(* Logix 5000 project; controller R400_500_XLS vendor 1 type 14 code 216 rev 31.11; software revision 31.01; part 7 of 32 *)
(* tags used below, declared in another part *)
   Abort1 : DINT;   // Not Used
   Abort2 : SINT;
   CURRENT_CYCLE : DINT;
   CycExcBuffer : UDT_CYCLE;
   CycleSequence : UDT_CYCLE_SEQUENCE;
   Drain_RcvryTnk_with_Sump : DINT;   // 0 = Close Recovery Tank Drain Valve 1 = Open Recovery Tank Drain Valve
   DrnSmp : DINT;
   DRYING : DINT;   // Drying id number
   F1rinse : DINT;   // Not Used
   F2rinse : DINT;   // Not Used
   F3rinse : DINT;   // Not Used
   FC65_Enabled_signal : BOOL;   // Enables the treatment evaluation
   FC65_Treatment_counter : DINT;   // Treatment counter
   Fill_Sump : DINT;
   FINALRINSE_1 : DINT;   // Final rinse 1 id number
   FINALRINSE_9 : DINT;   // Final rinse 9 id number
   HeatSmp : DINT;
   Inj_Time : SINT;   // Time based chemical injection steps
   M : DINT[5];   // Memory Bits
   ONS_FC13 : DINT;
   ONS_FC65 : DINT;
   OPR_16_TreatPrint_Ptr : DINT;
   PREWASH_1 : DINT;   // Pre-wash 1 id number
   PREWASH_2 : DINT;   // Pre-wash 2 id number
   PREWASH_3 : DINT;   // Pre-wash 3 id number
   PREWASH_4 : DINT;   // Pre-wash 4 id number
   printCycleParameters : STRING[2];
   PWHeat : SINT;
   Rcvry_Tnk_Tmp : REAL;   // Water Temperature of the Heat Recovery Tank
   RINSE_1 : DINT;   // Rinse 1 id number
   RINSE_2 : DINT;   // Rinse 2 id number
   RINSE_3 : DINT;   // Rinse 3 id number
   RINSE_4 : DINT;   // Rinse 4 id number
   Run : DINT;
   sCRLF : STRING;
   sPrntArray : STRING[300];   // Printer String Array
   SumpWaterVolume : DINT;   // Sump Water Volume 0 =Low 1= High
   Tmr : TIMER[107];
   Trt_Drying : SINT;
   Trt_PrWsh : DINT;
   Trt_Rinse : DINT;   // Rinse steps
   Trt_Wsh : DINT;
   VENTING : DINT;   // Venting id number
   WASH_1 : DINT;   // Wash 1 id number
   WASH_2 : DINT;   // Wash 2 id number
   WASH_3 : DINT;   // Wash 3 id number
   WASH_4 : DINT;   // Wash 4 id number
   WASH_5 : DINT;   // Wash 5 id number
   CycleName : STRING[12];
   EnaDisPrinter : BOOL;   // Screen 80 Enable/Disable Printer button
   msg : BOOL[512];
   Msg_Abort : SINT;
   PrintIndex : DINT;
   Screen_Ctrl : DINT;   // PLC Screen Request
   sDateTime : STRING;   // String Date Time
   Tpb : DINT[11];
   TreatmentPtr : DINT;
   Unit : Hrdwre;   // Unit Configuration
(* MainProgram, continued *)

ROUTINE OPR_15_WSH_13_ABORT   (* ladder *)
// This module manage the abort sequence.
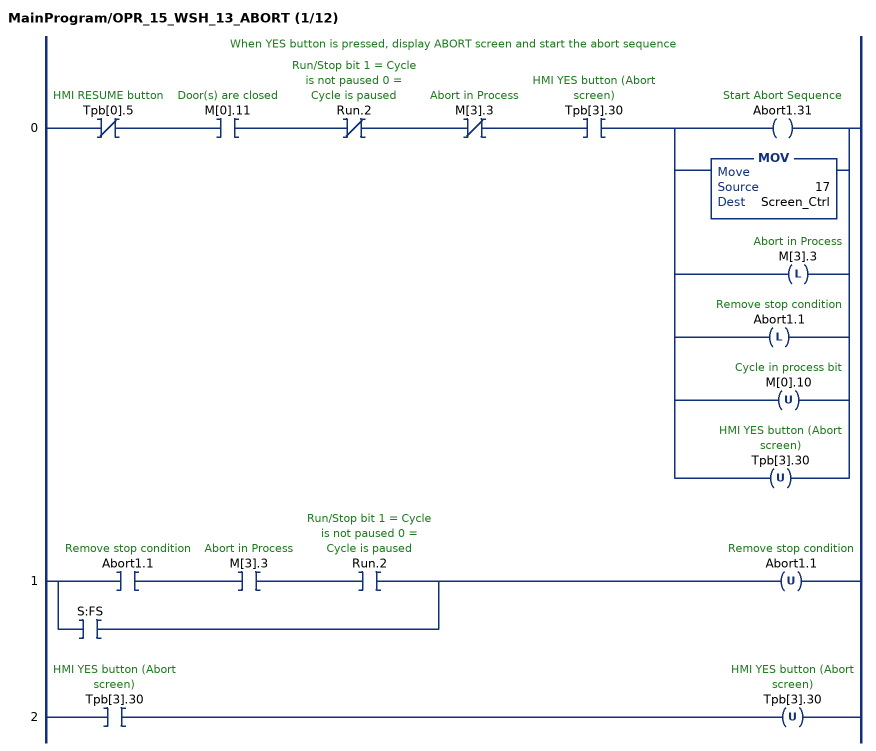
   // When YES button is pressed, display ABORT screen and start the abort sequence
   0: XIO(Tpb[0].5)XIC(M[0].11)XIO(Run.2)XIO(M[3].3)XIC(Tpb[3].30)[OTE(Abort1.31) ,MOV(17,Screen_Ctrl) ,OTL(M[3].3) ,OTL(Abort1.1) ,OTU(M[0].10) ,OTU(Tpb[3].30) ];
   1: [XIC(Abort1.1) XIC(M[3].3) XIC(Run.2) ,XIC(S:FS) ]OTU(Abort1.1);
   2: XIC(Tpb[3].30)OTU(Tpb[3].30);
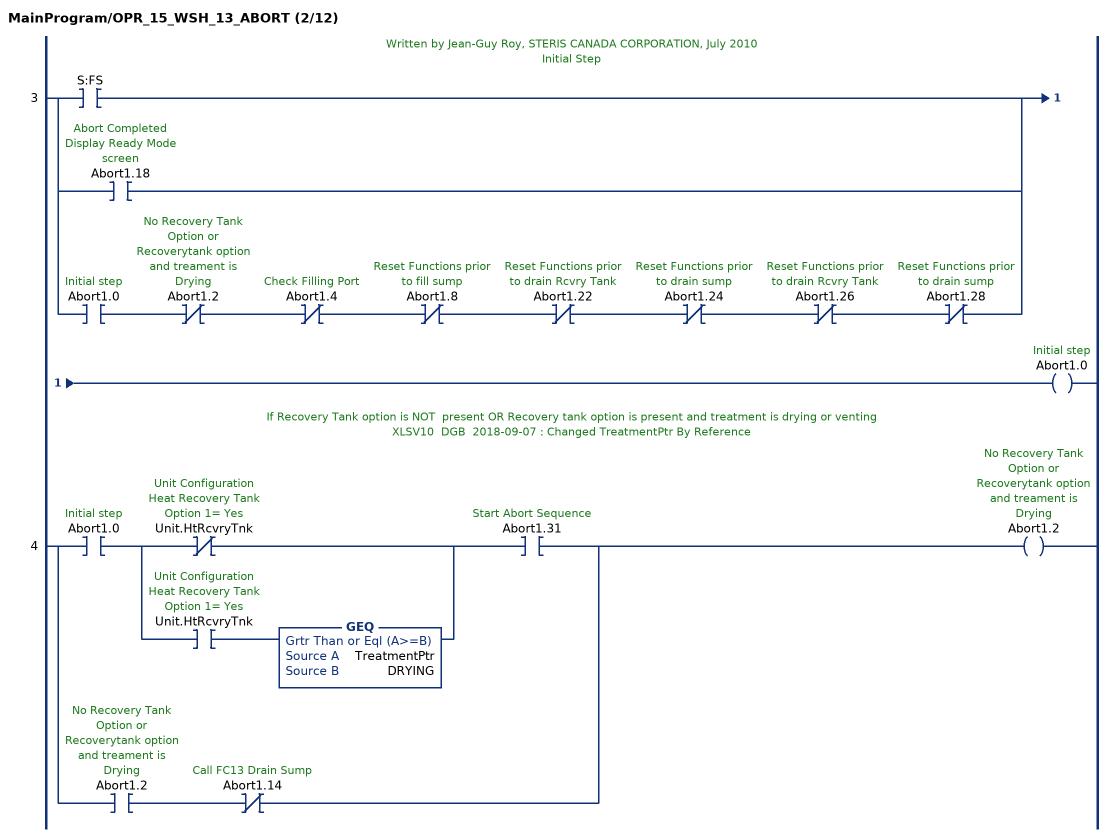
   // Written by Jean-Guy Roy, STERIS CANADA CORPORATION, July 2010
   // Initial Step
   3: [XIC(S:FS) ,XIC(Abort1.18) ,XIC(Abort1.0) XIO(Abort1.2) XIO(Abort1.4) XIO(Abort1.8) XIO(Abort1.22) XIO(Abort1.24) XIO(Abort1.26) XIO(Abort1.28) ]OTE(Abort1.0);
   // If Recovery Tank option is NOT  present OR Recovery tank option is present and treatment is drying or venting
   // XLSV10  DGB  2018-09-07 : Changed TreatmentPtr By Reference
   4: [XIC(Abort1.0) [XIO(Unit.HtRcvryTnk) ,XIC(Unit.HtRcvryTnk) GEQ(TreatmentPtr,DRYING) ] XIC(Abort1.31) ,XIC(Abort1.2) XIO(Abort1.14) ]OTE(Abort1.2);
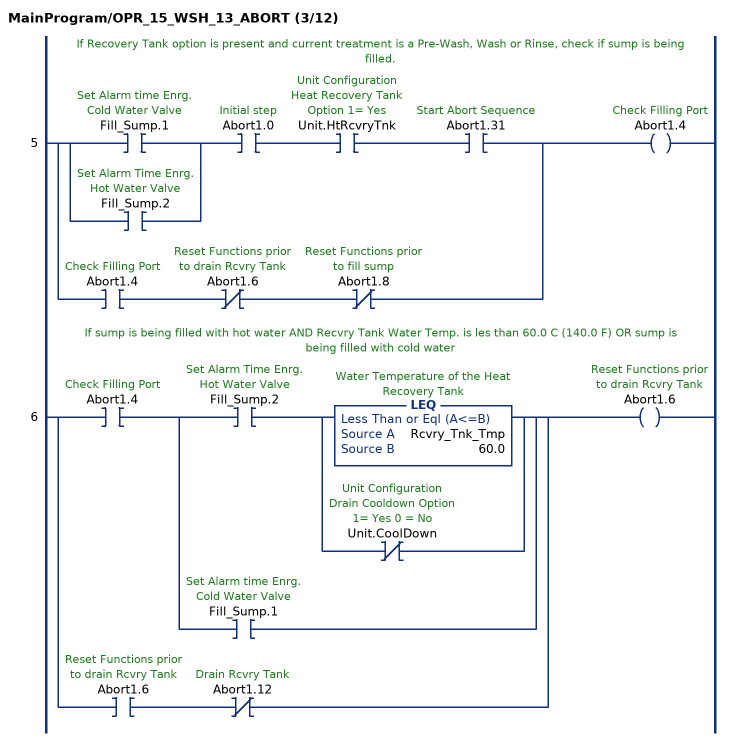
   // If Recovery Tank option is present and current treatment is a Pre-Wash, Wash or Rinse, check if sump is being filled.
   5: [[XIC(Fill_Sump.1) ,XIC(Fill_Sump.2) ] XIC(Abort1.0) XIC(Unit.HtRcvryTnk) XIC(Abort1.31) ,XIC(Abort1.4) XIO(Abort1.6) XIO(Abort1.8) ]OTE(Abort1.4);
   // If sump is being filled with hot water AND Recvry Tank Water Temp. is les than 60.0 C (140.0 F) OR sump is being filled with cold water
   6: [XIC(Abort1.4) [XIC(Fill_Sump.2) [LEQ(Rcvry_Tnk_Tmp,60.0) ,XIO(Unit.CoolDown) ] ,XIC(Fill_Sump.1) ] ,XIC(Abort1.6) XIO(Abort1.12) ]OTE(Abort1.6);
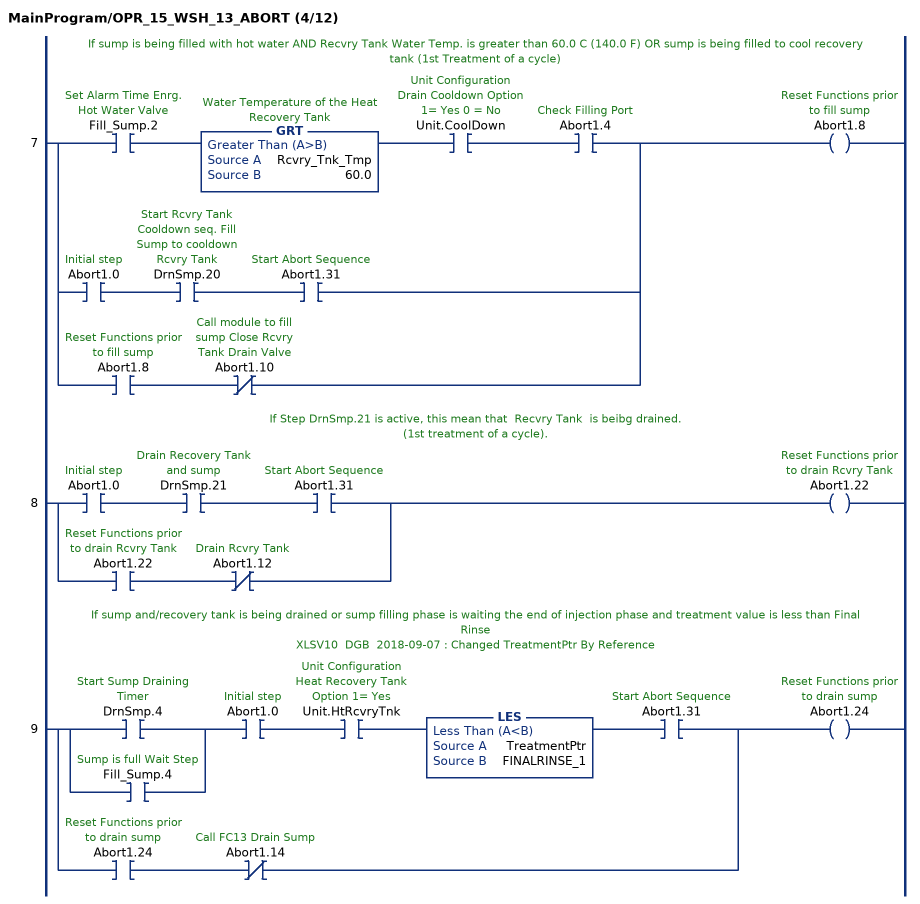
   // If sump is being filled with hot water AND Recvry Tank Water Temp. is greater than 60.0 C (140.0 F) OR sump is being filled to cool recovery tank (1st Treatment of a cycle)
   7: [[XIC(Fill_Sump.2) GRT(Rcvry_Tnk_Tmp,60.0) XIC(Unit.CoolDown) XIC(Abort1.4) ,XIC(Abort1.0) XIC(DrnSmp.20) XIC(Abort1.31) ] ,XIC(Abort1.8) XIO(Abort1.10) ]OTE(Abort1.8);
   // If Step DrnSmp.21 is active, this mean that  Recvry Tank  is beibg drained.
   //  (1st treatment of a cycle).
   8: [XIC(Abort1.0) XIC(DrnSmp.21) XIC(Abort1.31) ,XIC(Abort1.22) XIO(Abort1.12) ]OTE(Abort1.22);
   // If sump and/recovery tank is being drained or sump filling phase is waiting the end of injection phase and treatment value is less than Final Rinse
   // XLSV10  DGB  2018-09-07 : Changed TreatmentPtr By Reference
   9: [[XIC(DrnSmp.4) ,XIC(Fill_Sump.4) ] XIC(Abort1.0) XIC(Unit.HtRcvryTnk) LES(TreatmentPtr,FINALRINSE_1) XIC(Abort1.31) ,XIC(Abort1.24) XIO(Abort1.14) ]OTE(Abort1.24);
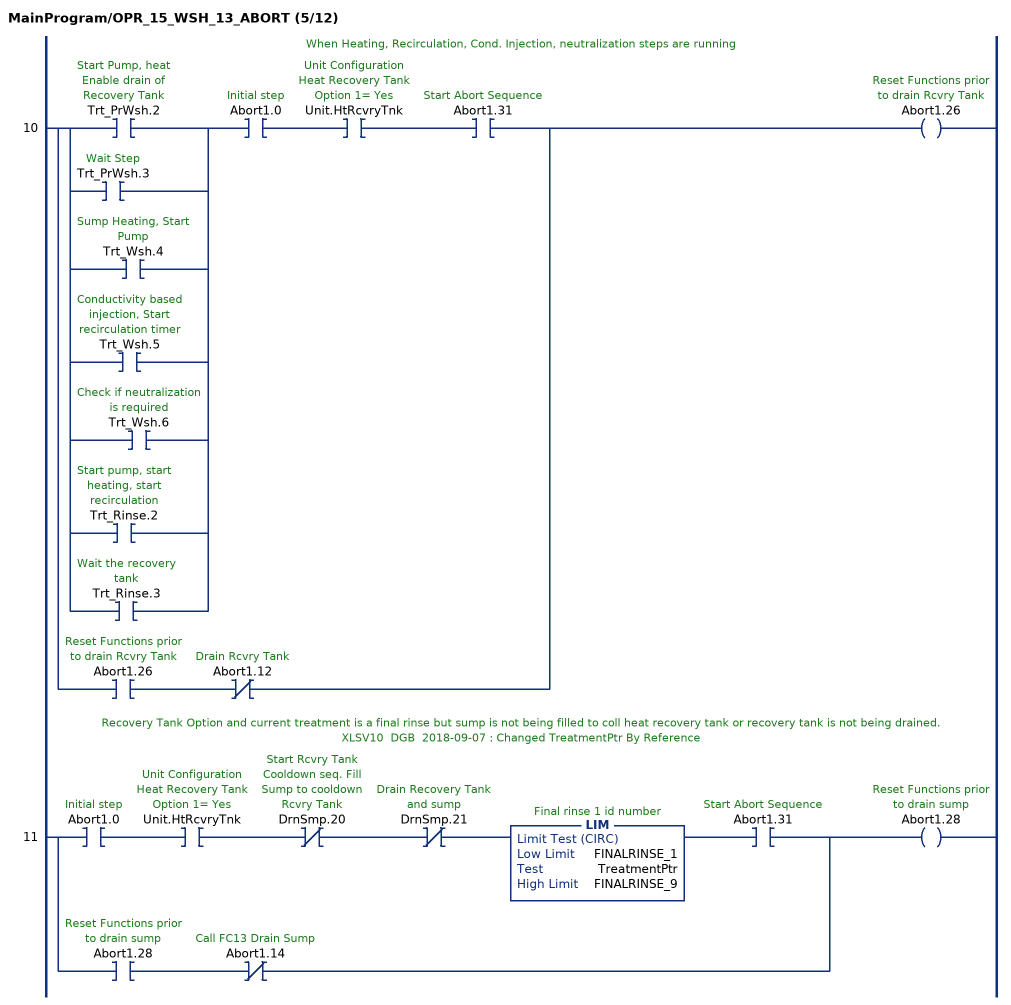
   // When Heating, Recirculation, Cond. Injection, neutralization steps are running
   10: [[XIC(Trt_PrWsh.2) ,XIC(Trt_PrWsh.3) ,XIC(Trt_Wsh.4) ,XIC(Trt_Wsh.5) ,XIC(Trt_Wsh.6) ,XIC(Trt_Rinse.2) ,XIC(Trt_Rinse.3) ] XIC(Abort1.0) XIC(Unit.HtRcvryTnk) XIC(Abort1.31) ,XIC(Abort1.26) XIO(Abort1.12) ]OTE(Abort1.26);
   // Recovery Tank Option and current treatment is a final rinse but sump is not being filled to coll heat recovery tank or recovery tank is not being drained.
   // XLSV10  DGB  2018-09-07 : Changed TreatmentPtr By Reference
   11: [XIC(Abort1.0) XIC(Unit.HtRcvryTnk) XIO(DrnSmp.20) XIO(DrnSmp.21) LIM(FINALRINSE_1,TreatmentPtr,FINALRINSE_9) XIC(Abort1.31) ,XIC(Abort1.28) XIO(Abort1.14) ]OTE(Abort1.28);
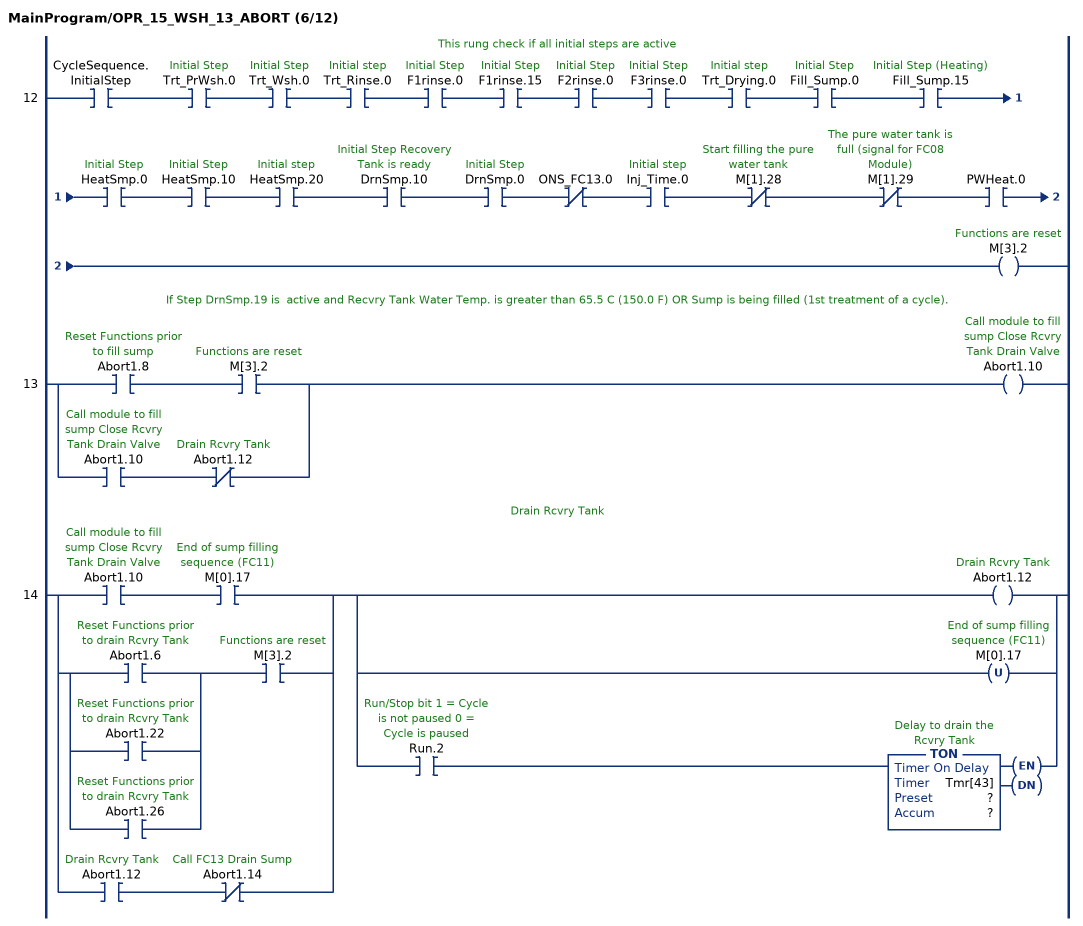
   // This rung check if all initial steps are active
   12: XIC(CycleSequence.InitialStep)XIC(Trt_PrWsh.0)XIC(Trt_Wsh.0)XIC(Trt_Rinse.0)XIC(F1rinse.0)XIC(F1rinse.15)XIC(F2rinse.0)XIC(F3rinse.0)XIC(Trt_Drying.0)XIC(Fill_Sump.0)XIC(Fill_Sump.15)XIC(HeatSmp.0)XIC(HeatSmp.10)XIC(HeatSmp.20)XIC(DrnSmp.10)XIC(DrnSmp.0)XIO(ONS_FC13.0)XIC(Inj_Time.0)XIO(M[1].28)XIO(M[1].29)XIC(PWHeat.0)OTE(M[3].2);
   // If Step DrnSmp.19 is  active and Recvry Tank Water Temp. is greater than 65.5 C (150.0 F) OR Sump is being filled (1st treatment of a cycle).
   13: [XIC(Abort1.8) XIC(M[3].2) ,XIC(Abort1.10) XIO(Abort1.12) ]OTE(Abort1.10);
   // Drain Rcvry Tank
   14: [XIC(Abort1.10) XIC(M[0].17) ,[XIC(Abort1.6) ,XIC(Abort1.22) ,XIC(Abort1.26) ] XIC(M[3].2) ,XIC(Abort1.12) XIO(Abort1.14) ][[OTE(Abort1.12) ,OTU(M[0].17) ] ,XIC(Run.2) TON(Tmr[43],?,?) ];
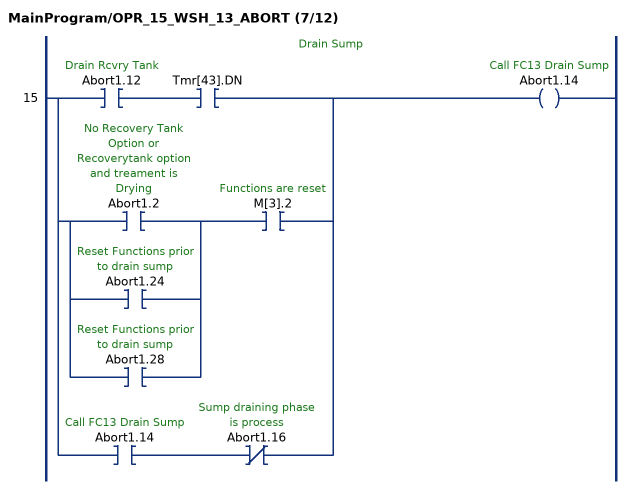
   // Drain Sump
   15: [XIC(Abort1.12) XIC(Tmr[43].DN) ,[XIC(Abort1.2) ,XIC(Abort1.24) ,XIC(Abort1.28) ] XIC(M[3].2) ,XIC(Abort1.14) XIO(Abort1.16) ]OTE(Abort1.14);
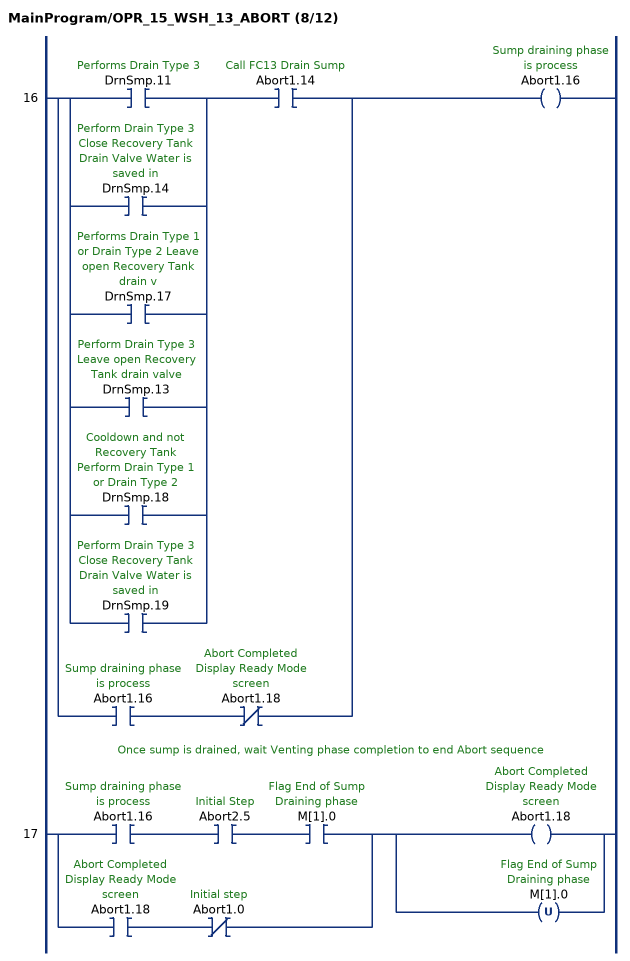
   16: [[XIC(DrnSmp.11) ,XIC(DrnSmp.14) ,XIC(DrnSmp.17) ,XIC(DrnSmp.13) ,XIC(DrnSmp.18) ,XIC(DrnSmp.19) ] XIC(Abort1.14) ,XIC(Abort1.16) XIO(Abort1.18) ]OTE(Abort1.16);
   // Once sump is drained, wait Venting phase completion to end Abort sequence
   17: [XIC(Abort1.16) XIC(Abort2.5) XIC(M[1].0) ,XIC(Abort1.18) XIO(Abort1.0) ][OTE(Abort1.18) ,OTU(M[1].0) ];
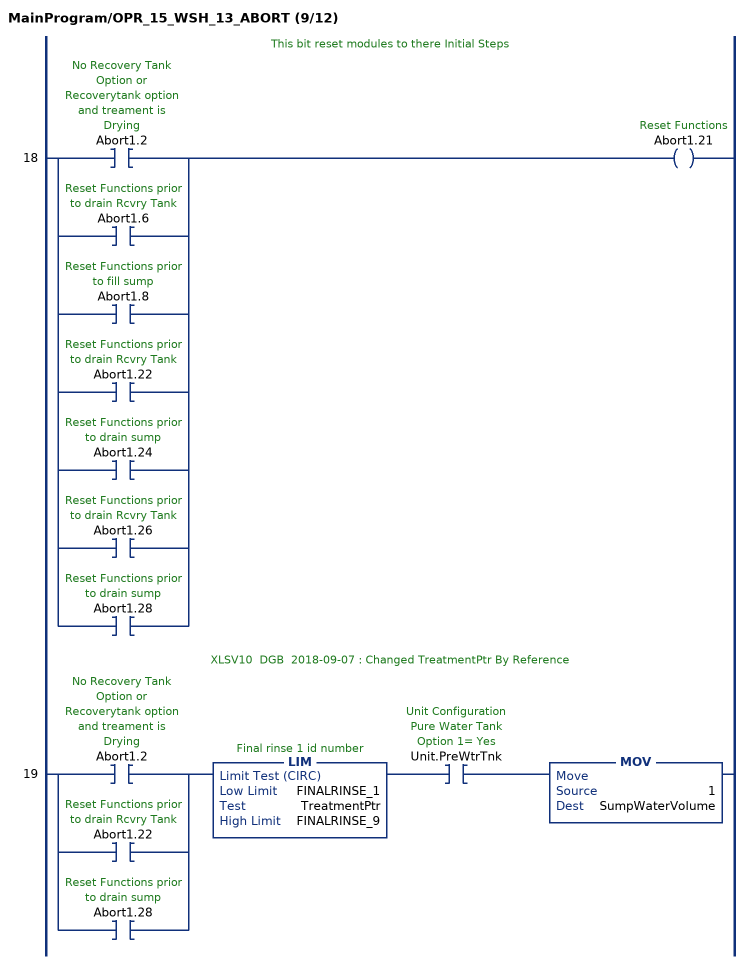
   // This bit reset modules to there Initial Steps
   18: [XIC(Abort1.2) ,XIC(Abort1.6) ,XIC(Abort1.8) ,XIC(Abort1.22) ,XIC(Abort1.24) ,XIC(Abort1.26) ,XIC(Abort1.28) ]OTE(Abort1.21);
   // XLSV10  DGB  2018-09-07 : Changed TreatmentPtr By Reference
   19: [XIC(Abort1.2) ,XIC(Abort1.22) ,XIC(Abort1.28) ]LIM(FINALRINSE_1,TreatmentPtr,FINALRINSE_9)XIC(Unit.PreWtrTnk)MOV(1,SumpWaterVolume);
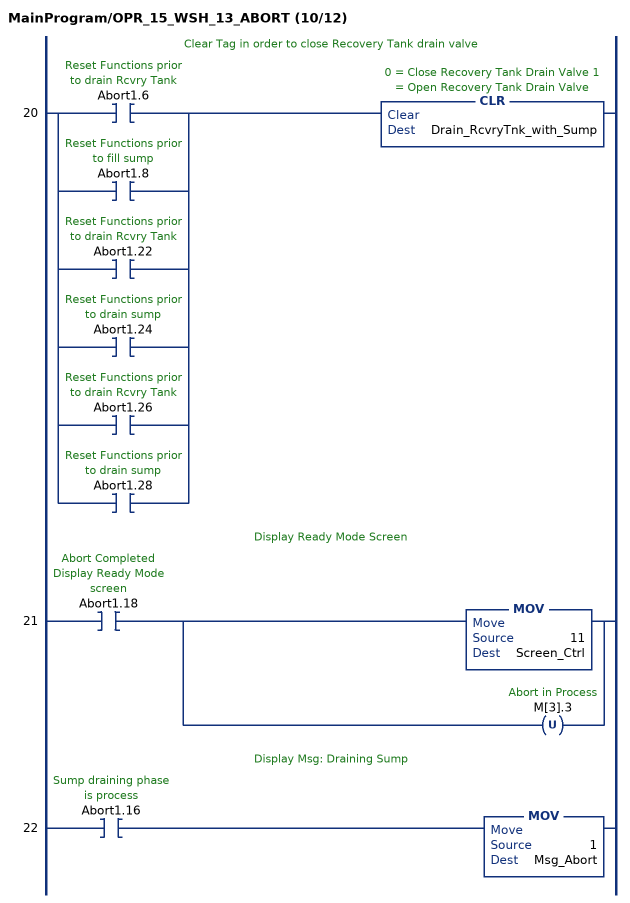
   // Clear Tag in order to close Recovery Tank drain valve
   20: [XIC(Abort1.6) ,XIC(Abort1.8) ,XIC(Abort1.22) ,XIC(Abort1.24) ,XIC(Abort1.26) ,XIC(Abort1.28) ]CLR(Drain_RcvryTnk_with_Sump);
   // Display Ready Mode Screen
   21: XIC(Abort1.18)[MOV(11,Screen_Ctrl) ,OTU(M[3].3) ];
   // Display Msg: Draining Sump
   22: XIC(Abort1.16)MOV(1,Msg_Abort);
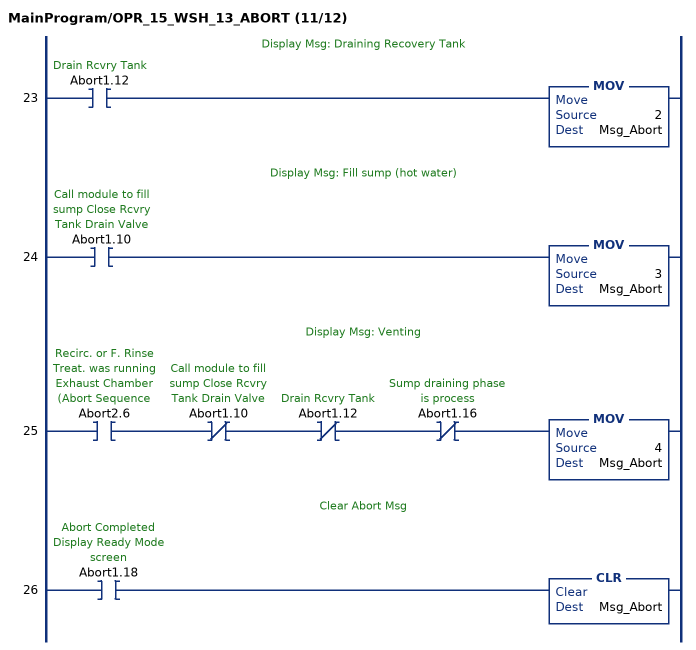
   // Display Msg: Draining Recovery Tank
   23: XIC(Abort1.12)MOV(2,Msg_Abort);
   // Display Msg: Fill sump (hot water)
   24: XIC(Abort1.10)MOV(3,Msg_Abort);
   // Display Msg: Venting
   25: XIC(Abort2.6)XIO(Abort1.10)XIO(Abort1.12)XIO(Abort1.16)MOV(4,Msg_Abort);
   // Clear Abort Msg
   26: XIC(Abort1.18)CLR(Msg_Abort);
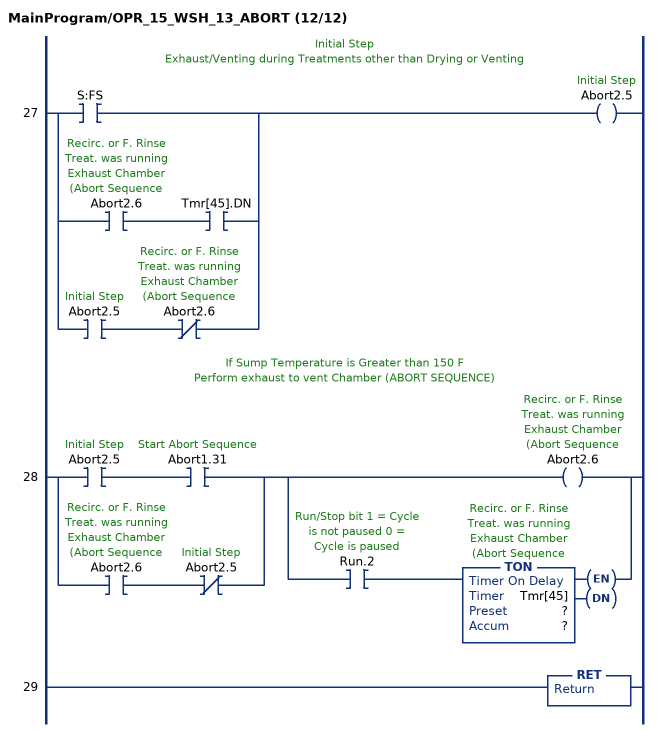
   // Initial Step
   // Exhaust/Venting during Treatments other than Drying or Venting
   27: [XIC(S:FS) ,XIC(Abort2.6) XIC(Tmr[45].DN) ,XIC(Abort2.5) XIO(Abort2.6) ]OTE(Abort2.5);
   // If Sump Temperature is Greater than 150 F
   // Perform exhaust to vent Chamber (ABORT SEQUENCE)
   28: [XIC(Abort2.5) XIC(Abort1.31) ,XIC(Abort2.6) XIO(Abort2.5) ][OTE(Abort2.6) ,XIC(Run.2) TON(Tmr[45],?,?) ];
   29: RET();
END_ROUTINE

ROUTINE OPR_16_PRINT_CYCLE_TREATMENTS   (* ladder *)
// This routines sends the treatment index to the WSH-38 requirement
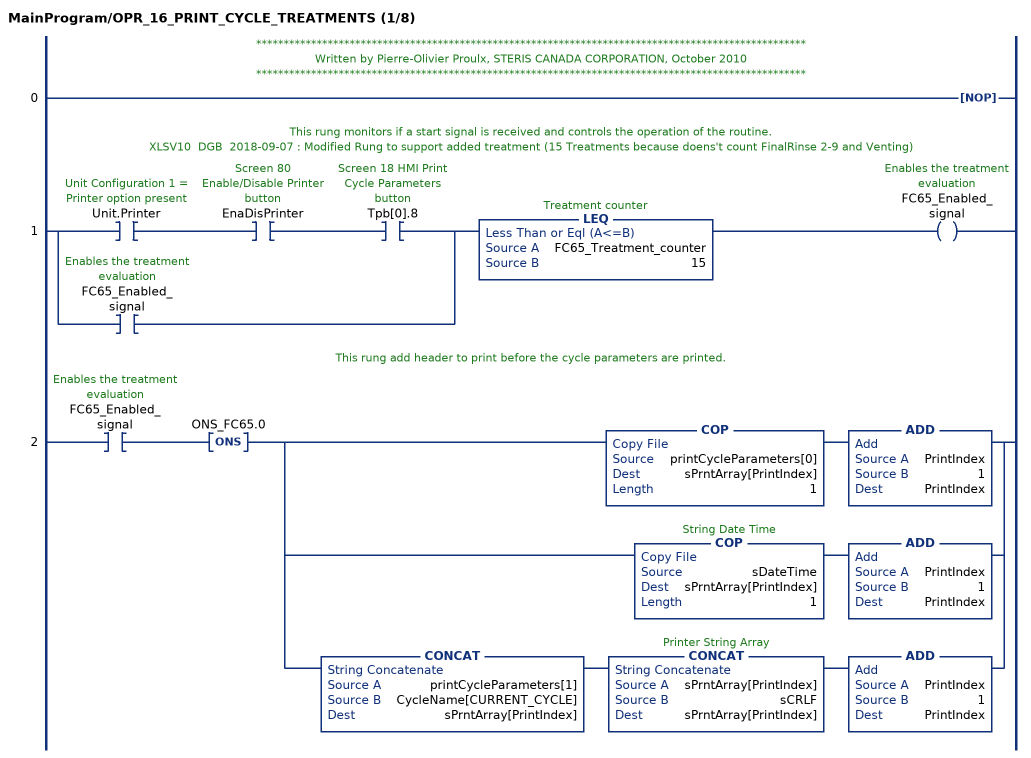
   // ****************************************************************************************************
   // Written by Pierre-Olivier Proulx, STERIS CANADA CORPORATION, October 2010
   // ****************************************************************************************************
   0: NOP();
   // This rung monitors if a start signal is received and controls the operation of the routine.
   // XLSV10  DGB  2018-09-07 : Modified Rung to support added treatment (15 Treatments because doens't count FinalRinse 2-9 and Venting)
   1: [XIC(Unit.Printer) XIC(EnaDisPrinter) XIC(Tpb[0].8) ,XIC(FC65_Enabled_signal) ]LEQ(FC65_Treatment_counter,15)OTE(FC65_Enabled_signal);
   // This rung add header to print before the cycle parameters are printed.
   2: XIC(FC65_Enabled_signal)ONS(ONS_FC65.0)[COP(printCycleParameters[0],sPrntArray[PrintIndex],1) ADD(PrintIndex,1,PrintIndex) ,COP(sDateTime,sPrntArray[PrintIndex],1) ADD(PrintIndex,1,PrintIndex) ,CONCAT(printCycleParameters[1],CycleName[CURRENT_CYCLE],sPrntArray[PrintIndex]) CONCAT(sPrntArray[PrintIndex],sCRLF,sPrntArray[PrintIndex]) ADD(PrintIndex,1,PrintIndex) ];
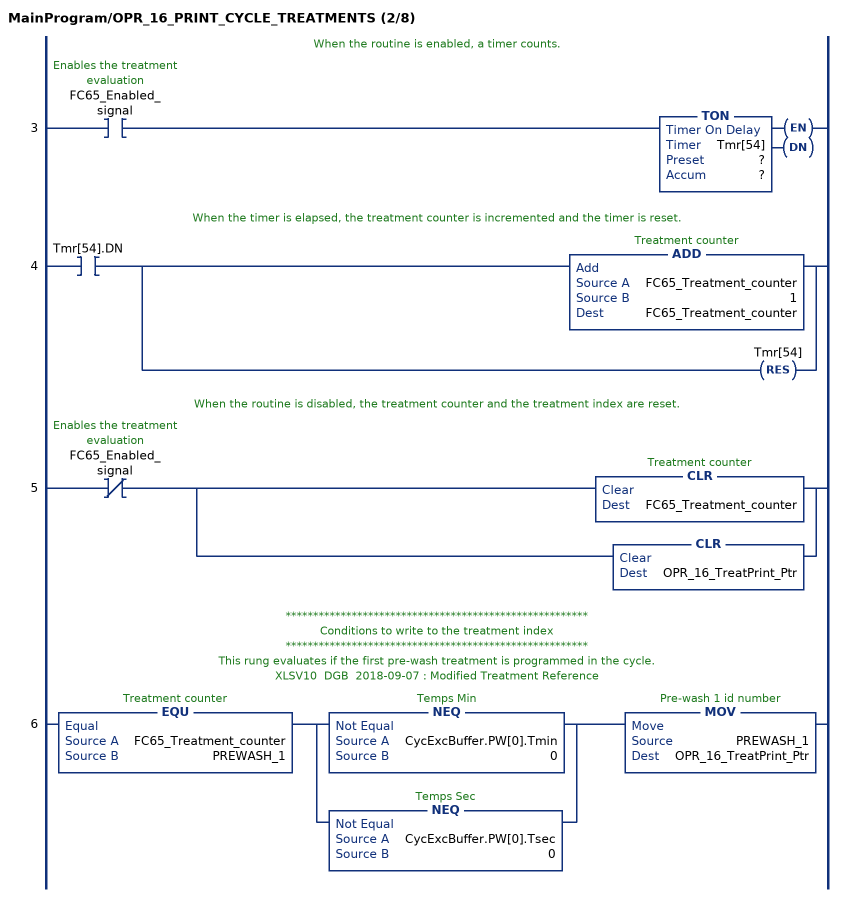
   // When the routine is enabled, a timer counts.
   3: XIC(FC65_Enabled_signal)TON(Tmr[54],?,?);
   // When the timer is elapsed, the treatment counter is incremented and the timer is reset.
   4: XIC(Tmr[54].DN)[ADD(FC65_Treatment_counter,1,FC65_Treatment_counter) ,RES(Tmr[54]) ];
   // When the routine is disabled, the treatment counter and the treatment index are reset.
   5: XIO(FC65_Enabled_signal)[CLR(FC65_Treatment_counter) ,CLR(OPR_16_TreatPrint_Ptr) ];
   // *******************************************************
   // Conditions to write to the treatment index
   // *******************************************************
   // This rung evaluates if the first pre-wash treatment is programmed in the cycle.
   // XLSV10  DGB  2018-09-07 : Modified Treatment Reference
   6: EQU(FC65_Treatment_counter,PREWASH_1)[NEQ(CycExcBuffer.PW[0].Tmin,0) ,NEQ(CycExcBuffer.PW[0].Tsec,0) ]MOV(PREWASH_1,OPR_16_TreatPrint_Ptr);
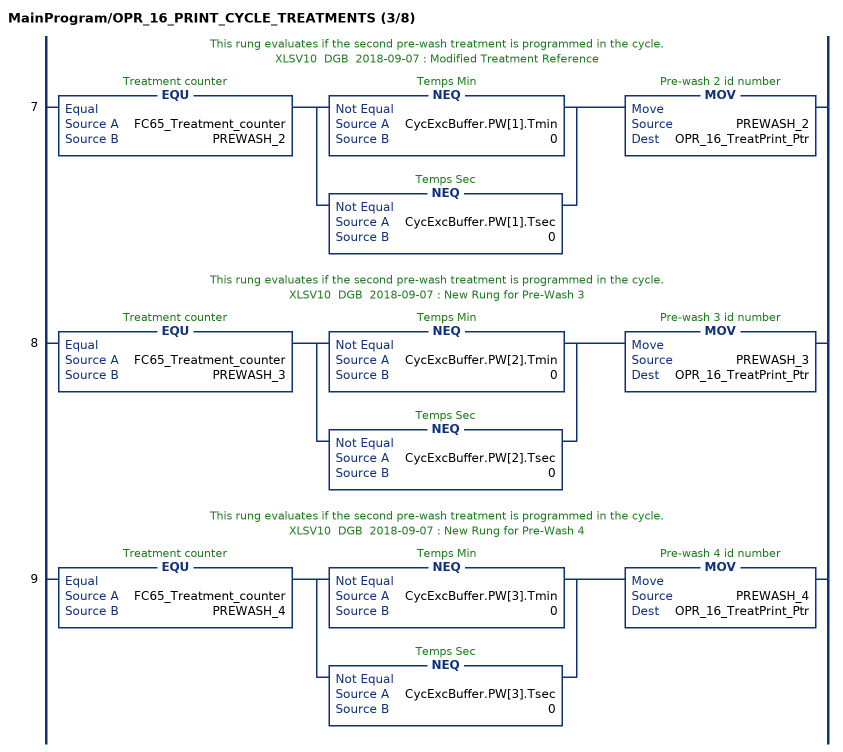
   // This rung evaluates if the second pre-wash treatment is programmed in the cycle.
   // XLSV10  DGB  2018-09-07 : Modified Treatment Reference
   7: EQU(FC65_Treatment_counter,PREWASH_2)[NEQ(CycExcBuffer.PW[1].Tmin,0) ,NEQ(CycExcBuffer.PW[1].Tsec,0) ]MOV(PREWASH_2,OPR_16_TreatPrint_Ptr);
   // This rung evaluates if the second pre-wash treatment is programmed in the cycle.
   // XLSV10  DGB  2018-09-07 : New Rung for Pre-Wash 3
   8: EQU(FC65_Treatment_counter,PREWASH_3)[NEQ(CycExcBuffer.PW[2].Tmin,0) ,NEQ(CycExcBuffer.PW[2].Tsec,0) ]MOV(PREWASH_3,OPR_16_TreatPrint_Ptr);
   // This rung evaluates if the second pre-wash treatment is programmed in the cycle.
   // XLSV10  DGB  2018-09-07 : New Rung for Pre-Wash 4
   9: EQU(FC65_Treatment_counter,PREWASH_4)[NEQ(CycExcBuffer.PW[3].Tmin,0) ,NEQ(CycExcBuffer.PW[3].Tsec,0) ]MOV(PREWASH_4,OPR_16_TreatPrint_Ptr);
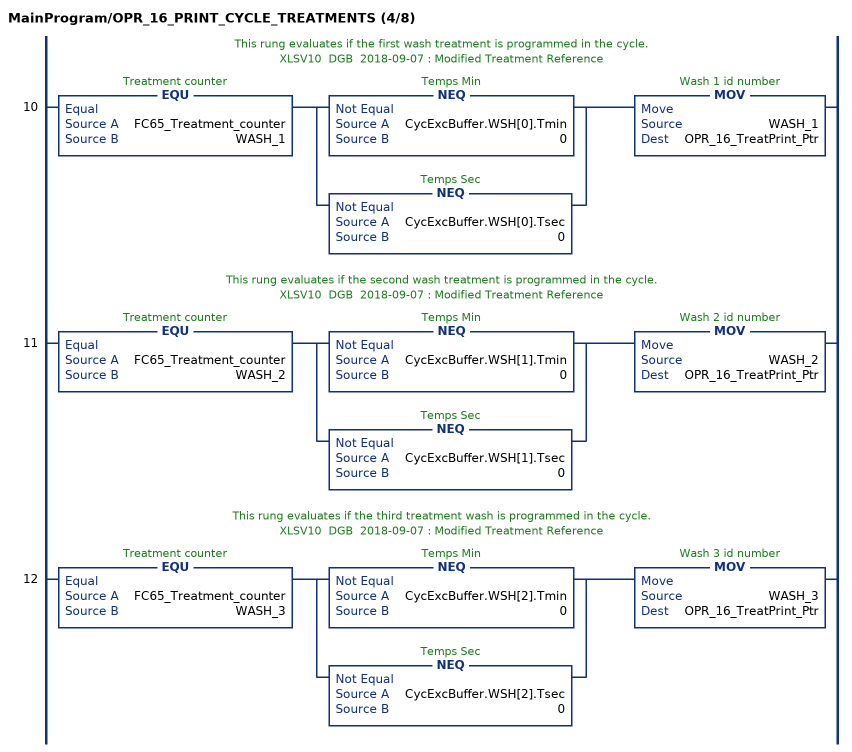
   // This rung evaluates if the first wash treatment is programmed in the cycle.
   // XLSV10  DGB  2018-09-07 : Modified Treatment Reference
   10: EQU(FC65_Treatment_counter,WASH_1)[NEQ(CycExcBuffer.WSH[0].Tmin,0) ,NEQ(CycExcBuffer.WSH[0].Tsec,0) ]MOV(WASH_1,OPR_16_TreatPrint_Ptr);
   // This rung evaluates if the second wash treatment is programmed in the cycle.
   // XLSV10  DGB  2018-09-07 : Modified Treatment Reference
   11: EQU(FC65_Treatment_counter,WASH_2)[NEQ(CycExcBuffer.WSH[1].Tmin,0) ,NEQ(CycExcBuffer.WSH[1].Tsec,0) ]MOV(WASH_2,OPR_16_TreatPrint_Ptr);
   // This rung evaluates if the third treatment wash is programmed in the cycle.
   // XLSV10  DGB  2018-09-07 : Modified Treatment Reference
   12: EQU(FC65_Treatment_counter,WASH_3)[NEQ(CycExcBuffer.WSH[2].Tmin,0) ,NEQ(CycExcBuffer.WSH[2].Tsec,0) ]MOV(WASH_3,OPR_16_TreatPrint_Ptr);
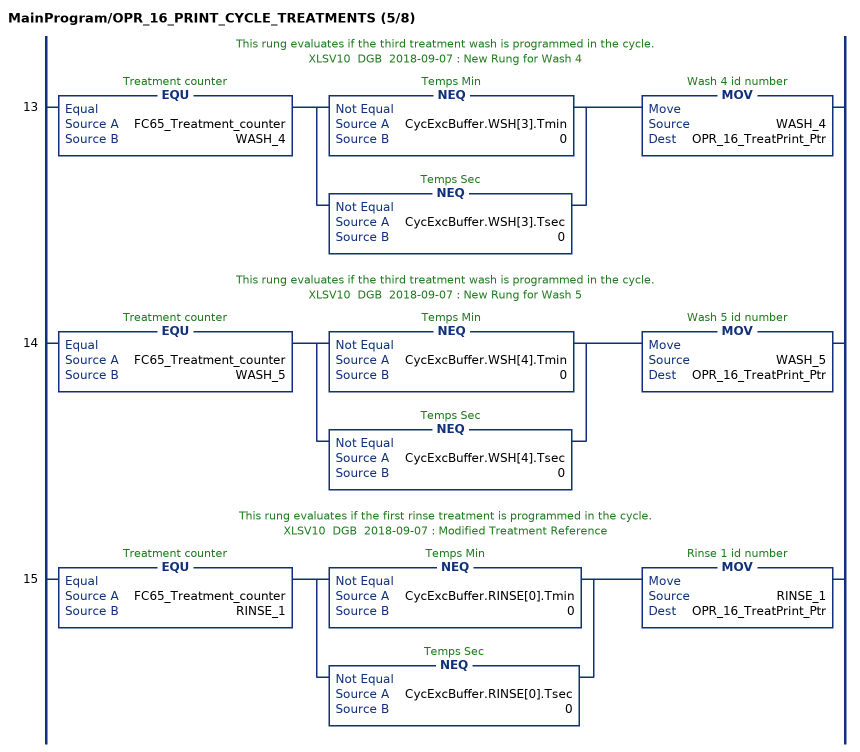
   // This rung evaluates if the third treatment wash is programmed in the cycle.
   // XLSV10  DGB  2018-09-07 : New Rung for Wash 4
   13: EQU(FC65_Treatment_counter,WASH_4)[NEQ(CycExcBuffer.WSH[3].Tmin,0) ,NEQ(CycExcBuffer.WSH[3].Tsec,0) ]MOV(WASH_4,OPR_16_TreatPrint_Ptr);
   // This rung evaluates if the third treatment wash is programmed in the cycle.
   // XLSV10  DGB  2018-09-07 : New Rung for Wash 5
   14: EQU(FC65_Treatment_counter,WASH_5)[NEQ(CycExcBuffer.WSH[4].Tmin,0) ,NEQ(CycExcBuffer.WSH[4].Tsec,0) ]MOV(WASH_5,OPR_16_TreatPrint_Ptr);
   // This rung evaluates if the first rinse treatment is programmed in the cycle.
   // XLSV10  DGB  2018-09-07 : Modified Treatment Reference
   15: EQU(FC65_Treatment_counter,RINSE_1)[NEQ(CycExcBuffer.RINSE[0].Tmin,0) ,NEQ(CycExcBuffer.RINSE[0].Tsec,0) ]MOV(RINSE_1,OPR_16_TreatPrint_Ptr);
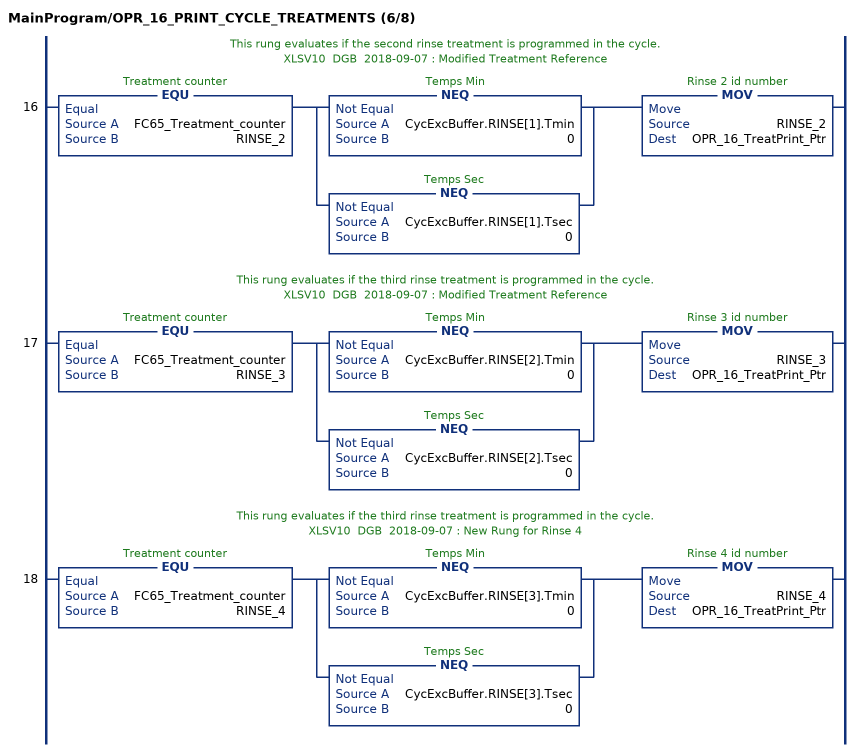
   // This rung evaluates if the second rinse treatment is programmed in the cycle.
   // XLSV10  DGB  2018-09-07 : Modified Treatment Reference
   16: EQU(FC65_Treatment_counter,RINSE_2)[NEQ(CycExcBuffer.RINSE[1].Tmin,0) ,NEQ(CycExcBuffer.RINSE[1].Tsec,0) ]MOV(RINSE_2,OPR_16_TreatPrint_Ptr);
   // This rung evaluates if the third rinse treatment is programmed in the cycle.
   // XLSV10  DGB  2018-09-07 : Modified Treatment Reference
   17: EQU(FC65_Treatment_counter,RINSE_3)[NEQ(CycExcBuffer.RINSE[2].Tmin,0) ,NEQ(CycExcBuffer.RINSE[2].Tsec,0) ]MOV(RINSE_3,OPR_16_TreatPrint_Ptr);
   // This rung evaluates if the third rinse treatment is programmed in the cycle.
   // XLSV10  DGB  2018-09-07 : New Rung for Rinse 4
   18: EQU(FC65_Treatment_counter,RINSE_4)[NEQ(CycExcBuffer.RINSE[3].Tmin,0) ,NEQ(CycExcBuffer.RINSE[3].Tsec,0) ]MOV(RINSE_4,OPR_16_TreatPrint_Ptr);
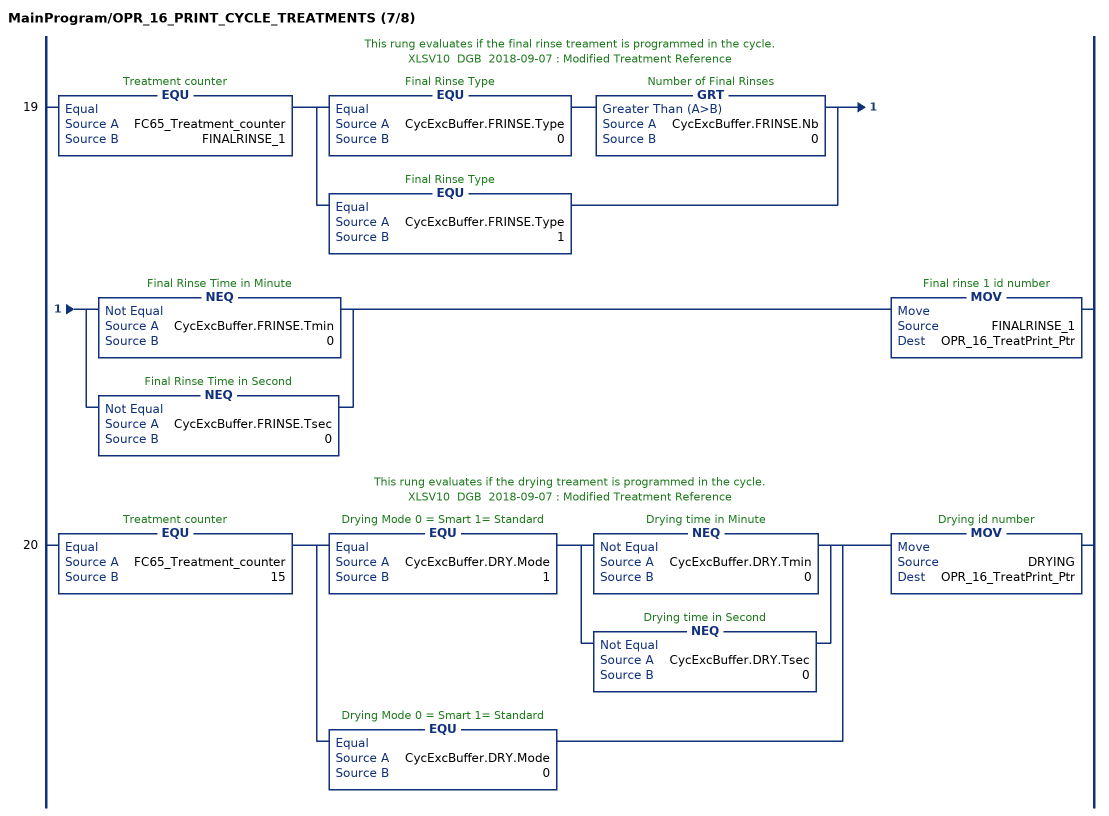
   // This rung evaluates if the final rinse treament is programmed in the cycle.
   // XLSV10  DGB  2018-09-07 : Modified Treatment Reference
   19: EQU(FC65_Treatment_counter,FINALRINSE_1)[EQU(CycExcBuffer.FRINSE.Type,0) GRT(CycExcBuffer.FRINSE.Nb,0) ,EQU(CycExcBuffer.FRINSE.Type,1) ][NEQ(CycExcBuffer.FRINSE.Tmin,0) ,NEQ(CycExcBuffer.FRINSE.Tsec,0) ]MOV(FINALRINSE_1,OPR_16_TreatPrint_Ptr);
   // This rung evaluates if the drying treament is programmed in the cycle.
   // XLSV10  DGB  2018-09-07 : Modified Treatment Reference
   20: EQU(FC65_Treatment_counter,15)[EQU(CycExcBuffer.DRY.Mode,1) [NEQ(CycExcBuffer.DRY.Tmin,0) ,NEQ(CycExcBuffer.DRY.Tsec,0) ] ,EQU(CycExcBuffer.DRY.Mode,0) ]MOV(DRYING,OPR_16_TreatPrint_Ptr);
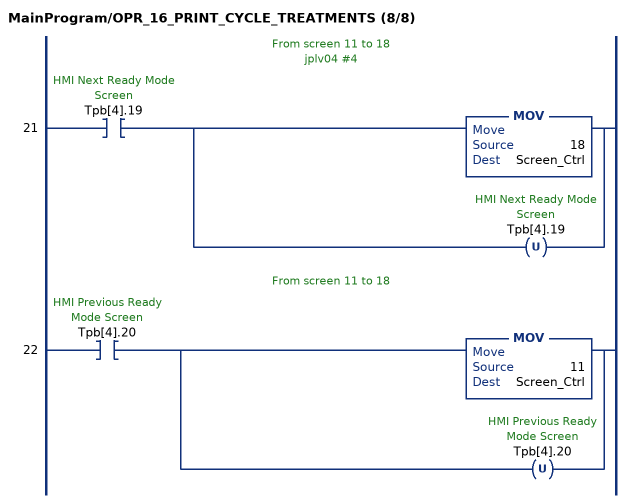
   // From screen 11 to 18
   // jplv04 #4
   21: XIC(Tpb[4].19)[MOV(18,Screen_Ctrl) ,OTU(Tpb[4].19) ];
   // From screen 11 to 18
   22: XIC(Tpb[4].20)[MOV(11,Screen_Ctrl) ,OTU(Tpb[4].20) ];
END_ROUTINE
